(* IEC 61131-3 sources: NachHouse_TST/ROOM_API_PILOT/getmem_test, 2 files *)

(* ---- 01_GETMEM_DATA.ST ---- *)
(* Fixed GETMEM test layout. All offsets are byte offsets from %R10000.

   0..3    ASCII "GMEM"
   4       format version = 1
   5       header size = 16
   6..7    payload size = 984, little-endian
   8..11   frame revision, little-endian
   12      pattern seed
   13..15  reserved, zero
   16..999 deterministic payload
*)

VAR_GLOBAL
    (* Raw memory read by: GETMEM:%R10000 1000 *)
    GetMemBuffer AT %R1000 : ARRAY[0..999] OF BYTE;

    (* Small public control/status surface. *)
    GetMemAddress     {PUBLIC_API} : STRING[16] := '%R1000';
    GetMemReadCommand {PUBLIC_API} : STRING[64] := 'GETMEM:%R1000 1000';
    GetMemLength      {PUBLIC_API} : UINT := 1000;
    GetMemRevision    {PUBLIC_API} : UDINT := 0;
    GetMemReady       {PUBLIC_API} : BOOL := FALSE;
    GetMemExecute     {PUBLIC_API} : BOOL := FALSE;
    GetMemSeed        {PUBLIC_API} : USINT := 0;

    GetMemInitialized : BOOL := FALSE;
END_VAR

FUNCTION GetMemBuildFrame : BOOL
VAR_INPUT
    Revision : UDINT;
    Seed     : USINT;
END_VAR
VAR
    i : UINT;
END_VAR

(* Fill the complete block first. *)
FOR i := 0 TO 999 DO
    GetMemBuffer[i] := UINT_TO_BYTE(i MOD 256) XOR USINT_TO_BYTE(Seed);
END_FOR;

(* Overwrite the first 16 bytes with a stable, easy-to-recognize header. *)
GetMemBuffer[0] := BYTE#16#47; (* G *)
GetMemBuffer[1] := BYTE#16#4D; (* M *)
GetMemBuffer[2] := BYTE#16#45; (* E *)
GetMemBuffer[3] := BYTE#16#4D; (* M *)
GetMemBuffer[4] := BYTE#1;
GetMemBuffer[5] := BYTE#16;
GetMemBuffer[6] := BYTE#16#D8; (* 984 = 16#03D8 *)
GetMemBuffer[7] := BYTE#16#03;
GetMemBuffer[8] := UDINT_TO_BYTE(Revision);
GetMemBuffer[9] := UDINT_TO_BYTE(SHR(Revision, 8));
GetMemBuffer[10] := UDINT_TO_BYTE(SHR(Revision, 16));
GetMemBuffer[11] := UDINT_TO_BYTE(SHR(Revision, 24));
GetMemBuffer[12] := USINT_TO_BYTE(Seed);
GetMemBuffer[13] := BYTE#0;
GetMemBuffer[14] := BYTE#0;
GetMemBuffer[15] := BYTE#0;

GetMemBuildFrame := TRUE;
END_FUNCTION

(* ---- prgMain.ST ---- *)
PROGRAM prgMain
VAR
    nextRevision : UDINT;
    nextSeed     : USINT;
END_VAR

(* Build a known first frame after program start. *)
IF NOT GetMemInitialized THEN
    GetMemReady := FALSE;
    GetMemBuildFrame(Revision := 1, Seed := 0);
    GetMemSeed := 0;
    GetMemRevision := 1; (* Commit is published only after the buffer is complete. *)
    GetMemReady := TRUE;
    GetMemInitialized := TRUE;
END_IF;

(* A SET of GetMemExecute=TRUE creates a visibly different test frame. *)
IF GetMemExecute THEN
    GetMemReady := FALSE;
    nextRevision := GetMemRevision + 1;
    nextSeed := GetMemSeed + 1;
    GetMemBuildFrame(Revision := nextRevision, Seed := nextSeed);
    GetMemSeed := nextSeed;
    GetMemRevision := nextRevision; (* Commit last. *)
    GetMemReady := TRUE;
    GetMemExecute := FALSE;
END_IF;
END_PROGRAM
